(* Logix 5000 project; controller CIP vendor 1 type 14 code 106 rev 20.12; software revision 20.06; part 8 of 13 *)
(* tags used below, declared in another part *)
   MOA_OFF : DINT[10];
   MOA_ON : DINT[10];
   PV_Output_Status : INT[10];
   PV_Output_Status_IND : INT[10,16];
   PV_Status_Bit : BOOL;
   Time_Date : DINT[20];
(* MainProgram, continued *)

ROUTINE _10_PV_STATUS   (* ladder *)
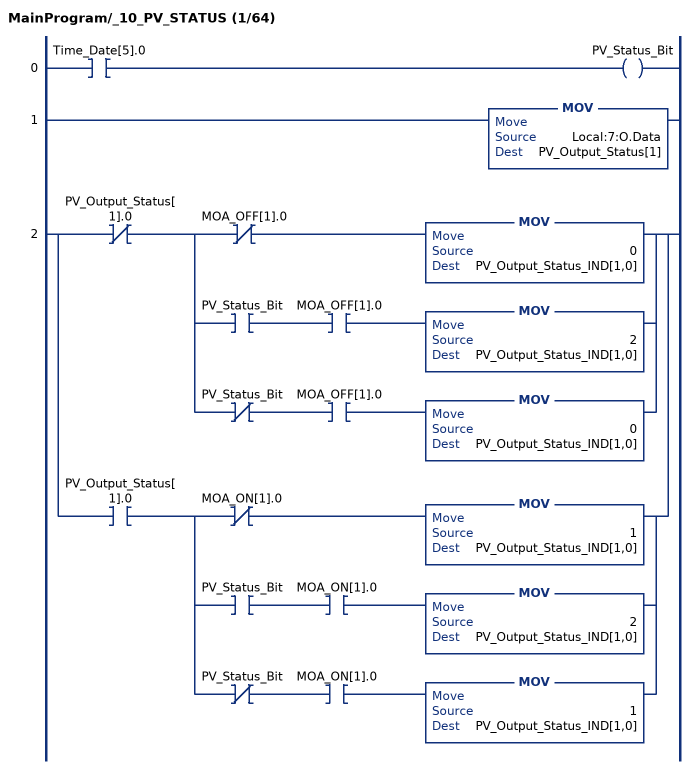
   0: XIC(Time_Date[5].0)OTE(PV_Status_Bit);
   1: MOV(Local:7:O.Data,PV_Output_Status[1]);
   2: [XIO(PV_Output_Status[1].0) [XIO(MOA_OFF[1].0) MOV(0,PV_Output_Status_IND[1,0]) ,XIC(PV_Status_Bit) XIC(MOA_OFF[1].0) MOV(2,PV_Output_Status_IND[1,0]) ,XIO(PV_Status_Bit) XIC(MOA_OFF[1].0) MOV(0,PV_Output_Status_IND[1,0]) ] ,XIC(PV_Output_Status[1].0) [XIO(MOA_ON[1].0) MOV(1,PV_Output_Status_IND[1,0]) ,XIC(PV_Status_Bit) XIC(MOA_ON[1].0) MOV(2,PV_Output_Status_IND[1,0]) ,XIO(PV_Status_Bit) XIC(MOA_ON[1].0) MOV(1,PV_Output_Status_IND[1,0]) ] ];
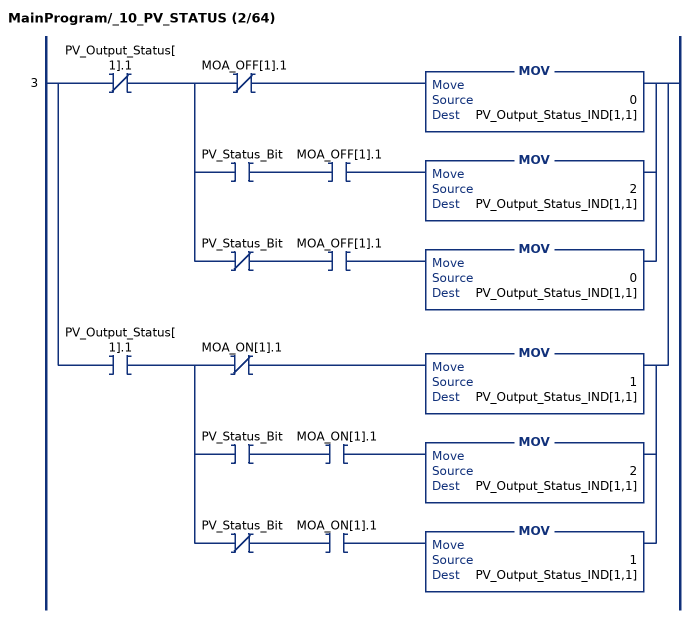
   3: [XIO(PV_Output_Status[1].1) [XIO(MOA_OFF[1].1) MOV(0,PV_Output_Status_IND[1,1]) ,XIC(PV_Status_Bit) XIC(MOA_OFF[1].1) MOV(2,PV_Output_Status_IND[1,1]) ,XIO(PV_Status_Bit) XIC(MOA_OFF[1].1) MOV(0,PV_Output_Status_IND[1,1]) ] ,XIC(PV_Output_Status[1].1) [XIO(MOA_ON[1].1) MOV(1,PV_Output_Status_IND[1,1]) ,XIC(PV_Status_Bit) XIC(MOA_ON[1].1) MOV(2,PV_Output_Status_IND[1,1]) ,XIO(PV_Status_Bit) XIC(MOA_ON[1].1) MOV(1,PV_Output_Status_IND[1,1]) ] ];
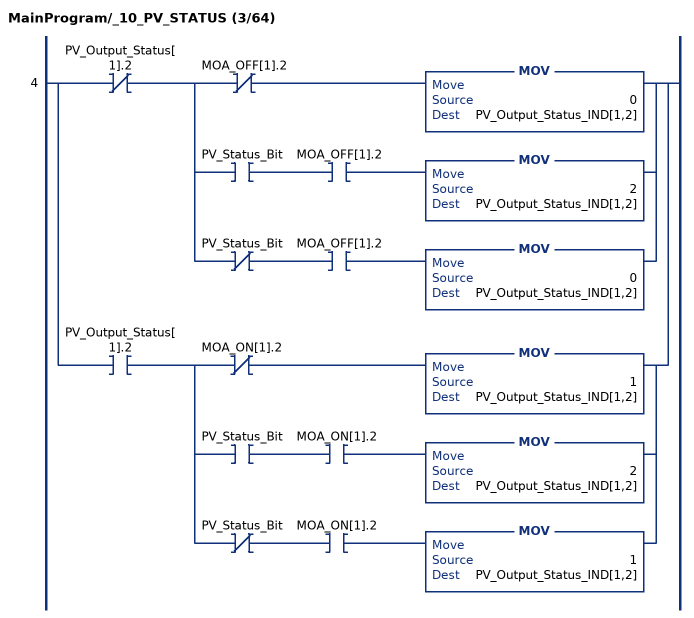
   4: [XIO(PV_Output_Status[1].2) [XIO(MOA_OFF[1].2) MOV(0,PV_Output_Status_IND[1,2]) ,XIC(PV_Status_Bit) XIC(MOA_OFF[1].2) MOV(2,PV_Output_Status_IND[1,2]) ,XIO(PV_Status_Bit) XIC(MOA_OFF[1].2) MOV(0,PV_Output_Status_IND[1,2]) ] ,XIC(PV_Output_Status[1].2) [XIO(MOA_ON[1].2) MOV(1,PV_Output_Status_IND[1,2]) ,XIC(PV_Status_Bit) XIC(MOA_ON[1].2) MOV(2,PV_Output_Status_IND[1,2]) ,XIO(PV_Status_Bit) XIC(MOA_ON[1].2) MOV(1,PV_Output_Status_IND[1,2]) ] ];
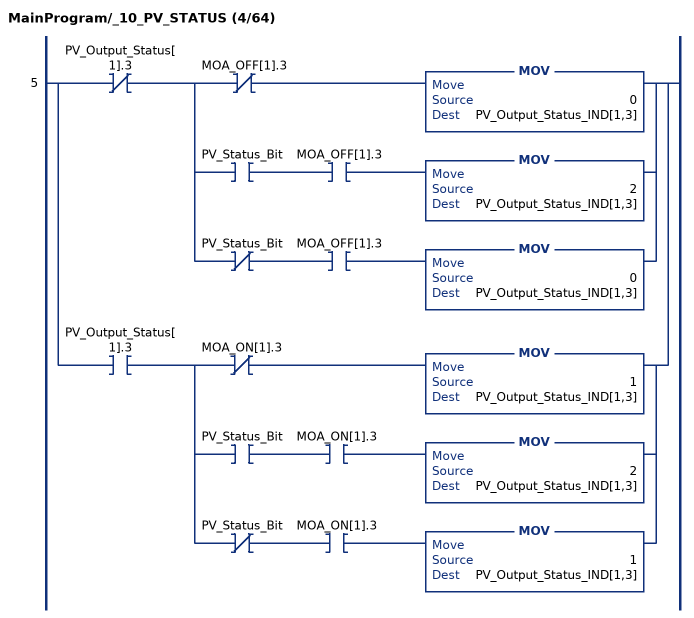
   5: [XIO(PV_Output_Status[1].3) [XIO(MOA_OFF[1].3) MOV(0,PV_Output_Status_IND[1,3]) ,XIC(PV_Status_Bit) XIC(MOA_OFF[1].3) MOV(2,PV_Output_Status_IND[1,3]) ,XIO(PV_Status_Bit) XIC(MOA_OFF[1].3) MOV(0,PV_Output_Status_IND[1,3]) ] ,XIC(PV_Output_Status[1].3) [XIO(MOA_ON[1].3) MOV(1,PV_Output_Status_IND[1,3]) ,XIC(PV_Status_Bit) XIC(MOA_ON[1].3) MOV(2,PV_Output_Status_IND[1,3]) ,XIO(PV_Status_Bit) XIC(MOA_ON[1].3) MOV(1,PV_Output_Status_IND[1,3]) ] ];
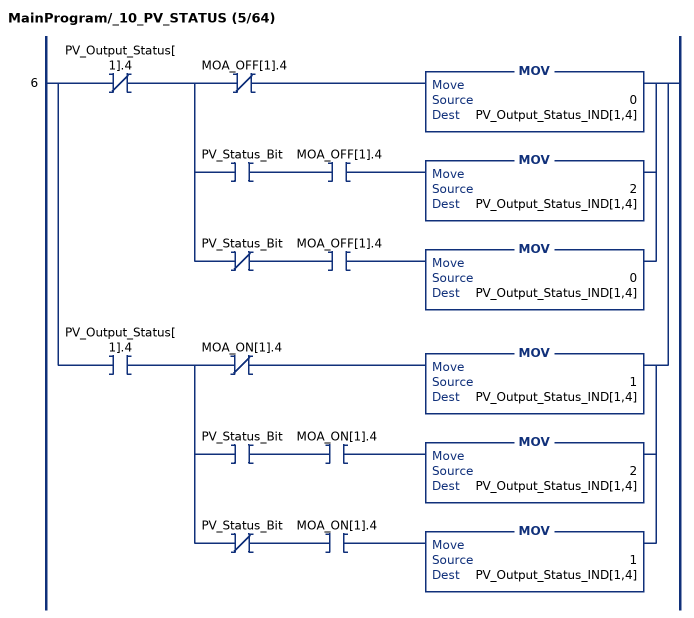
   6: [XIO(PV_Output_Status[1].4) [XIO(MOA_OFF[1].4) MOV(0,PV_Output_Status_IND[1,4]) ,XIC(PV_Status_Bit) XIC(MOA_OFF[1].4) MOV(2,PV_Output_Status_IND[1,4]) ,XIO(PV_Status_Bit) XIC(MOA_OFF[1].4) MOV(0,PV_Output_Status_IND[1,4]) ] ,XIC(PV_Output_Status[1].4) [XIO(MOA_ON[1].4) MOV(1,PV_Output_Status_IND[1,4]) ,XIC(PV_Status_Bit) XIC(MOA_ON[1].4) MOV(2,PV_Output_Status_IND[1,4]) ,XIO(PV_Status_Bit) XIC(MOA_ON[1].4) MOV(1,PV_Output_Status_IND[1,4]) ] ];
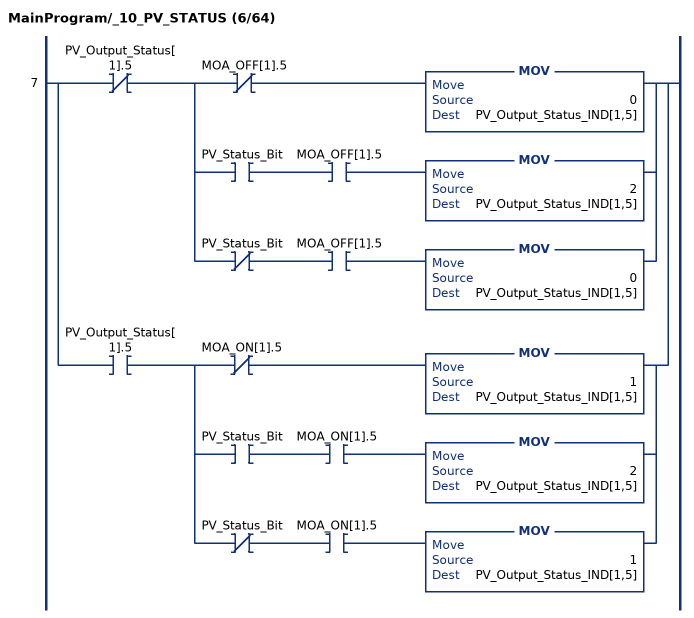
   7: [XIO(PV_Output_Status[1].5) [XIO(MOA_OFF[1].5) MOV(0,PV_Output_Status_IND[1,5]) ,XIC(PV_Status_Bit) XIC(MOA_OFF[1].5) MOV(2,PV_Output_Status_IND[1,5]) ,XIO(PV_Status_Bit) XIC(MOA_OFF[1].5) MOV(0,PV_Output_Status_IND[1,5]) ] ,XIC(PV_Output_Status[1].5) [XIO(MOA_ON[1].5) MOV(1,PV_Output_Status_IND[1,5]) ,XIC(PV_Status_Bit) XIC(MOA_ON[1].5) MOV(2,PV_Output_Status_IND[1,5]) ,XIO(PV_Status_Bit) XIC(MOA_ON[1].5) MOV(1,PV_Output_Status_IND[1,5]) ] ];
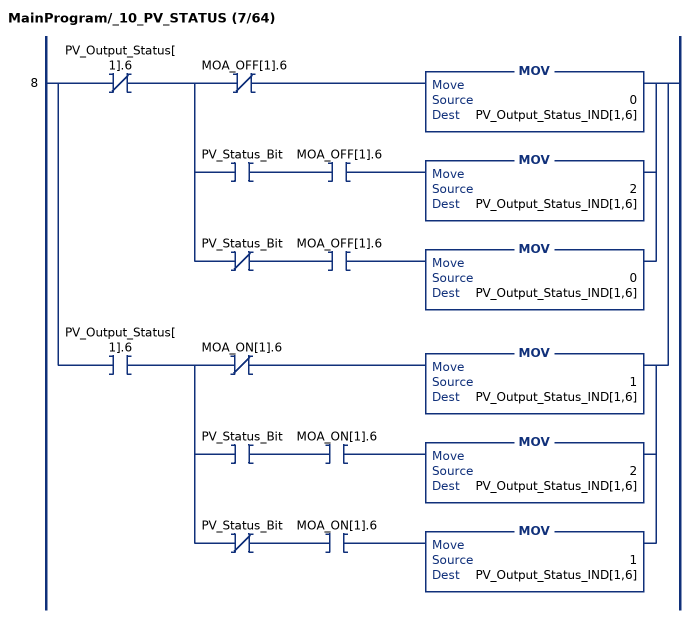
   8: [XIO(PV_Output_Status[1].6) [XIO(MOA_OFF[1].6) MOV(0,PV_Output_Status_IND[1,6]) ,XIC(PV_Status_Bit) XIC(MOA_OFF[1].6) MOV(2,PV_Output_Status_IND[1,6]) ,XIO(PV_Status_Bit) XIC(MOA_OFF[1].6) MOV(0,PV_Output_Status_IND[1,6]) ] ,XIC(PV_Output_Status[1].6) [XIO(MOA_ON[1].6) MOV(1,PV_Output_Status_IND[1,6]) ,XIC(PV_Status_Bit) XIC(MOA_ON[1].6) MOV(2,PV_Output_Status_IND[1,6]) ,XIO(PV_Status_Bit) XIC(MOA_ON[1].6) MOV(1,PV_Output_Status_IND[1,6]) ] ];
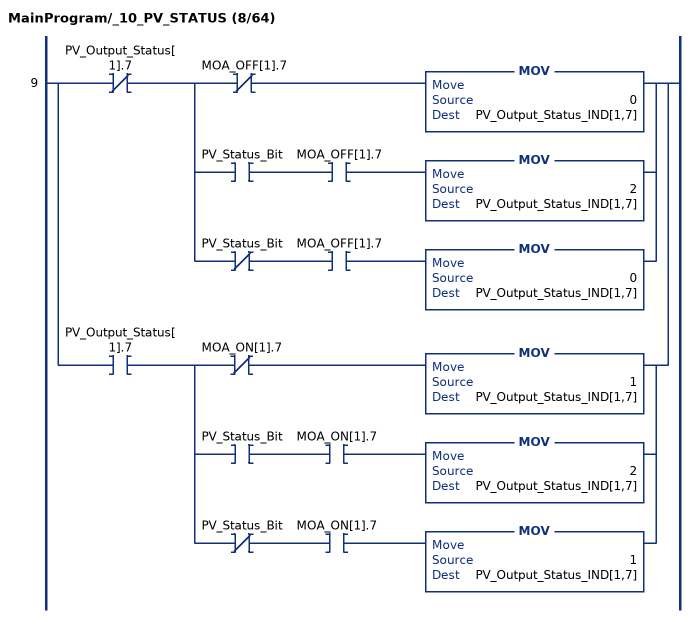
   9: [XIO(PV_Output_Status[1].7) [XIO(MOA_OFF[1].7) MOV(0,PV_Output_Status_IND[1,7]) ,XIC(PV_Status_Bit) XIC(MOA_OFF[1].7) MOV(2,PV_Output_Status_IND[1,7]) ,XIO(PV_Status_Bit) XIC(MOA_OFF[1].7) MOV(0,PV_Output_Status_IND[1,7]) ] ,XIC(PV_Output_Status[1].7) [XIO(MOA_ON[1].7) MOV(1,PV_Output_Status_IND[1,7]) ,XIC(PV_Status_Bit) XIC(MOA_ON[1].7) MOV(2,PV_Output_Status_IND[1,7]) ,XIO(PV_Status_Bit) XIC(MOA_ON[1].7) MOV(1,PV_Output_Status_IND[1,7]) ] ];
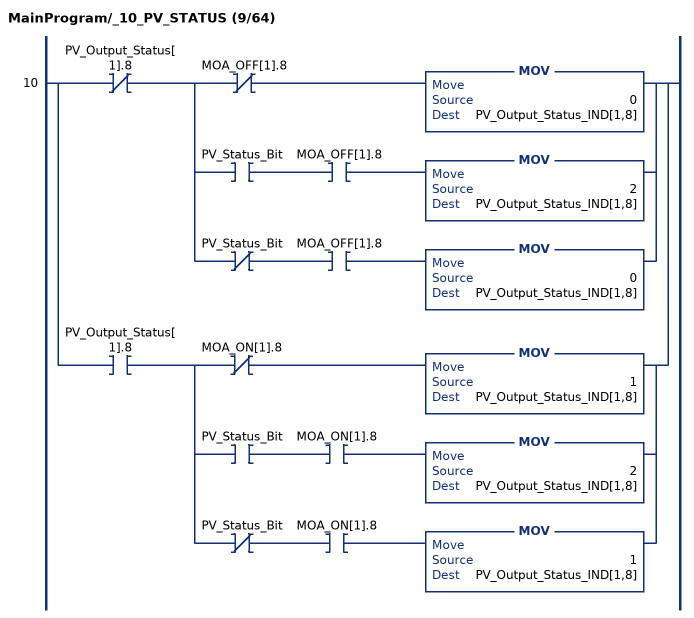
   10: [XIO(PV_Output_Status[1].8) [XIO(MOA_OFF[1].8) MOV(0,PV_Output_Status_IND[1,8]) ,XIC(PV_Status_Bit) XIC(MOA_OFF[1].8) MOV(2,PV_Output_Status_IND[1,8]) ,XIO(PV_Status_Bit) XIC(MOA_OFF[1].8) MOV(0,PV_Output_Status_IND[1,8]) ] ,XIC(PV_Output_Status[1].8) [XIO(MOA_ON[1].8) MOV(1,PV_Output_Status_IND[1,8]) ,XIC(PV_Status_Bit) XIC(MOA_ON[1].8) MOV(2,PV_Output_Status_IND[1,8]) ,XIO(PV_Status_Bit) XIC(MOA_ON[1].8) MOV(1,PV_Output_Status_IND[1,8]) ] ];
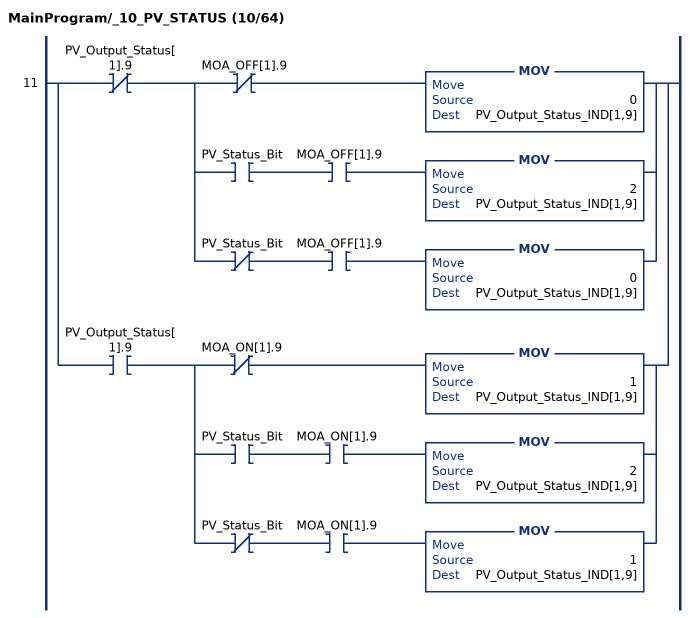
   11: [XIO(PV_Output_Status[1].9) [XIO(MOA_OFF[1].9) MOV(0,PV_Output_Status_IND[1,9]) ,XIC(PV_Status_Bit) XIC(MOA_OFF[1].9) MOV(2,PV_Output_Status_IND[1,9]) ,XIO(PV_Status_Bit) XIC(MOA_OFF[1].9) MOV(0,PV_Output_Status_IND[1,9]) ] ,XIC(PV_Output_Status[1].9) [XIO(MOA_ON[1].9) MOV(1,PV_Output_Status_IND[1,9]) ,XIC(PV_Status_Bit) XIC(MOA_ON[1].9) MOV(2,PV_Output_Status_IND[1,9]) ,XIO(PV_Status_Bit) XIC(MOA_ON[1].9) MOV(1,PV_Output_Status_IND[1,9]) ] ];
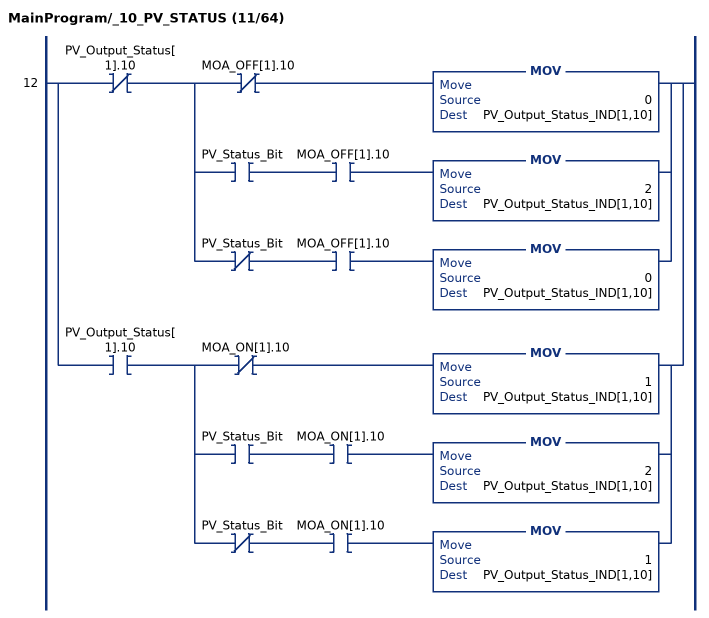
   12: [XIO(PV_Output_Status[1].10) [XIO(MOA_OFF[1].10) MOV(0,PV_Output_Status_IND[1,10]) ,XIC(PV_Status_Bit) XIC(MOA_OFF[1].10) MOV(2,PV_Output_Status_IND[1,10]) ,XIO(PV_Status_Bit) XIC(MOA_OFF[1].10) MOV(0,PV_Output_Status_IND[1,10]) ] ,XIC(PV_Output_Status[1].10) [XIO(MOA_ON[1].10) MOV(1,PV_Output_Status_IND[1,10]) ,XIC(PV_Status_Bit) XIC(MOA_ON[1].10) MOV(2,PV_Output_Status_IND[1,10]) ,XIO(PV_Status_Bit) XIC(MOA_ON[1].10) MOV(1,PV_Output_Status_IND[1,10]) ] ];
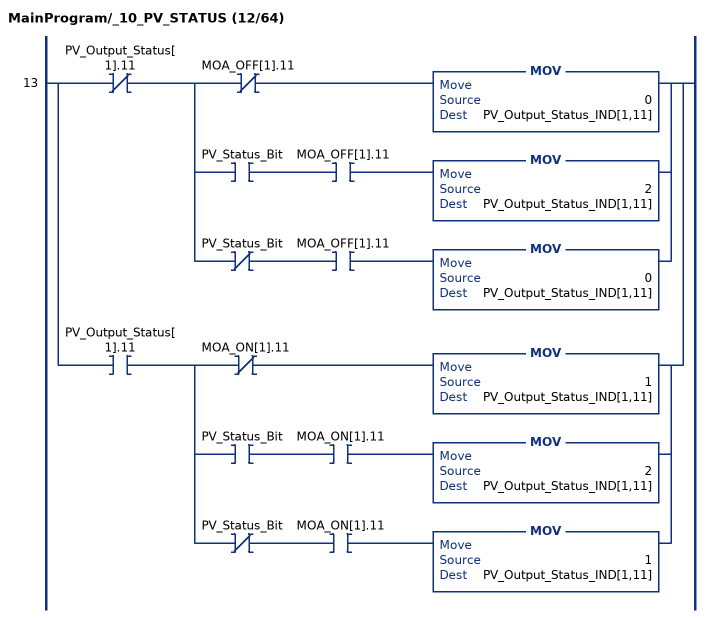
   13: [XIO(PV_Output_Status[1].11) [XIO(MOA_OFF[1].11) MOV(0,PV_Output_Status_IND[1,11]) ,XIC(PV_Status_Bit) XIC(MOA_OFF[1].11) MOV(2,PV_Output_Status_IND[1,11]) ,XIO(PV_Status_Bit) XIC(MOA_OFF[1].11) MOV(0,PV_Output_Status_IND[1,11]) ] ,XIC(PV_Output_Status[1].11) [XIO(MOA_ON[1].11) MOV(1,PV_Output_Status_IND[1,11]) ,XIC(PV_Status_Bit) XIC(MOA_ON[1].11) MOV(2,PV_Output_Status_IND[1,11]) ,XIO(PV_Status_Bit) XIC(MOA_ON[1].11) MOV(1,PV_Output_Status_IND[1,11]) ] ];
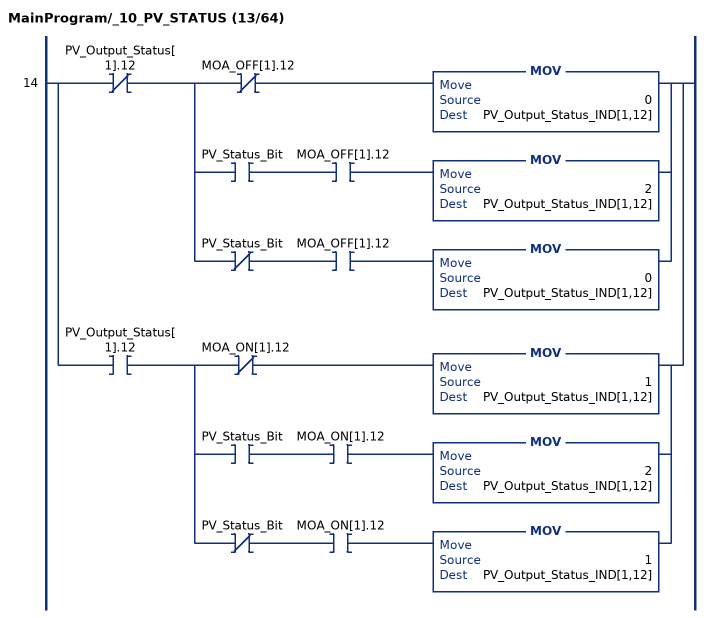
   14: [XIO(PV_Output_Status[1].12) [XIO(MOA_OFF[1].12) MOV(0,PV_Output_Status_IND[1,12]) ,XIC(PV_Status_Bit) XIC(MOA_OFF[1].12) MOV(2,PV_Output_Status_IND[1,12]) ,XIO(PV_Status_Bit) XIC(MOA_OFF[1].12) MOV(0,PV_Output_Status_IND[1,12]) ] ,XIC(PV_Output_Status[1].12) [XIO(MOA_ON[1].12) MOV(1,PV_Output_Status_IND[1,12]) ,XIC(PV_Status_Bit) XIC(MOA_ON[1].12) MOV(2,PV_Output_Status_IND[1,12]) ,XIO(PV_Status_Bit) XIC(MOA_ON[1].12) MOV(1,PV_Output_Status_IND[1,12]) ] ];
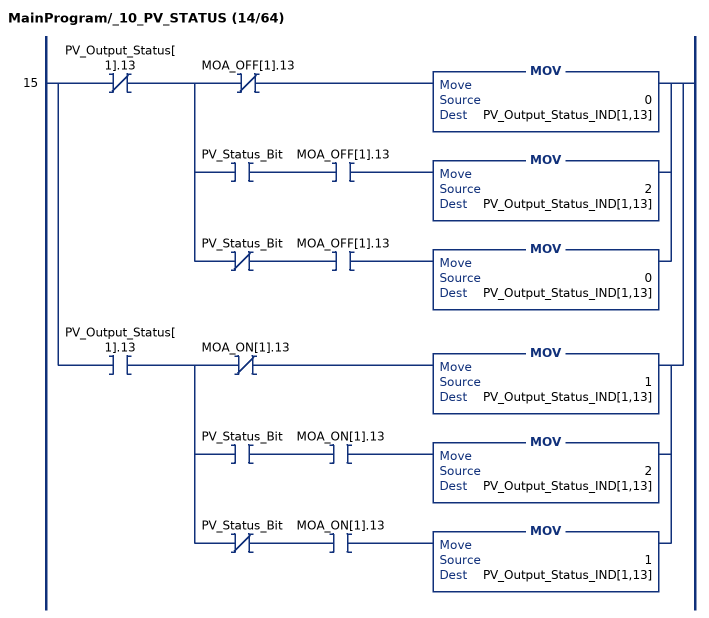
   15: [XIO(PV_Output_Status[1].13) [XIO(MOA_OFF[1].13) MOV(0,PV_Output_Status_IND[1,13]) ,XIC(PV_Status_Bit) XIC(MOA_OFF[1].13) MOV(2,PV_Output_Status_IND[1,13]) ,XIO(PV_Status_Bit) XIC(MOA_OFF[1].13) MOV(0,PV_Output_Status_IND[1,13]) ] ,XIC(PV_Output_Status[1].13) [XIO(MOA_ON[1].13) MOV(1,PV_Output_Status_IND[1,13]) ,XIC(PV_Status_Bit) XIC(MOA_ON[1].13) MOV(2,PV_Output_Status_IND[1,13]) ,XIO(PV_Status_Bit) XIC(MOA_ON[1].13) MOV(1,PV_Output_Status_IND[1,13]) ] ];
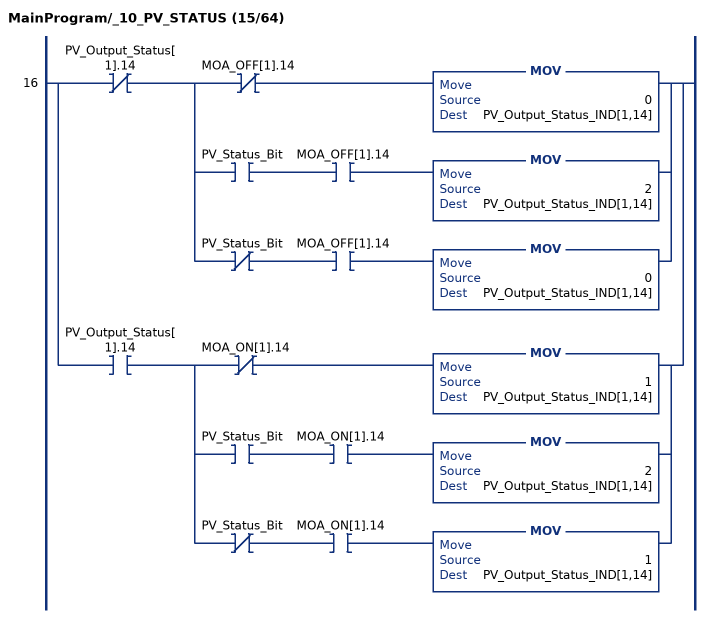
   16: [XIO(PV_Output_Status[1].14) [XIO(MOA_OFF[1].14) MOV(0,PV_Output_Status_IND[1,14]) ,XIC(PV_Status_Bit) XIC(MOA_OFF[1].14) MOV(2,PV_Output_Status_IND[1,14]) ,XIO(PV_Status_Bit) XIC(MOA_OFF[1].14) MOV(0,PV_Output_Status_IND[1,14]) ] ,XIC(PV_Output_Status[1].14) [XIO(MOA_ON[1].14) MOV(1,PV_Output_Status_IND[1,14]) ,XIC(PV_Status_Bit) XIC(MOA_ON[1].14) MOV(2,PV_Output_Status_IND[1,14]) ,XIO(PV_Status_Bit) XIC(MOA_ON[1].14) MOV(1,PV_Output_Status_IND[1,14]) ] ];
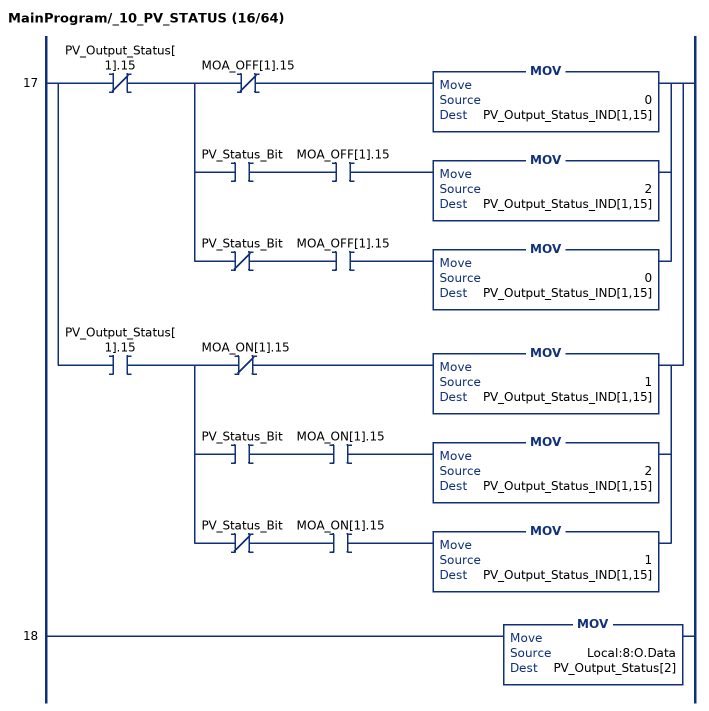
   17: [XIO(PV_Output_Status[1].15) [XIO(MOA_OFF[1].15) MOV(0,PV_Output_Status_IND[1,15]) ,XIC(PV_Status_Bit) XIC(MOA_OFF[1].15) MOV(2,PV_Output_Status_IND[1,15]) ,XIO(PV_Status_Bit) XIC(MOA_OFF[1].15) MOV(0,PV_Output_Status_IND[1,15]) ] ,XIC(PV_Output_Status[1].15) [XIO(MOA_ON[1].15) MOV(1,PV_Output_Status_IND[1,15]) ,XIC(PV_Status_Bit) XIC(MOA_ON[1].15) MOV(2,PV_Output_Status_IND[1,15]) ,XIO(PV_Status_Bit) XIC(MOA_ON[1].15) MOV(1,PV_Output_Status_IND[1,15]) ] ];
   18: MOV(Local:8:O.Data,PV_Output_Status[2]);
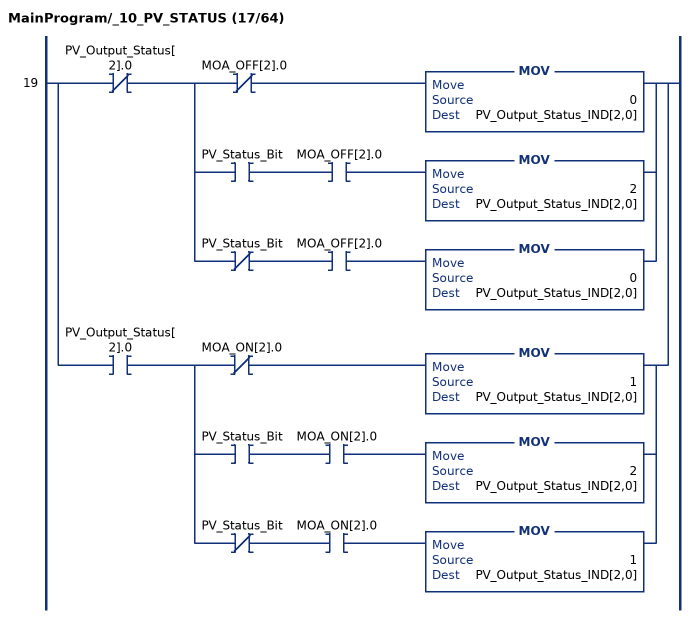
   19: [XIO(PV_Output_Status[2].0) [XIO(MOA_OFF[2].0) MOV(0,PV_Output_Status_IND[2,0]) ,XIC(PV_Status_Bit) XIC(MOA_OFF[2].0) MOV(2,PV_Output_Status_IND[2,0]) ,XIO(PV_Status_Bit) XIC(MOA_OFF[2].0) MOV(0,PV_Output_Status_IND[2,0]) ] ,XIC(PV_Output_Status[2].0) [XIO(MOA_ON[2].0) MOV(1,PV_Output_Status_IND[2,0]) ,XIC(PV_Status_Bit) XIC(MOA_ON[2].0) MOV(2,PV_Output_Status_IND[2,0]) ,XIO(PV_Status_Bit) XIC(MOA_ON[2].0) MOV(1,PV_Output_Status_IND[2,0]) ] ];
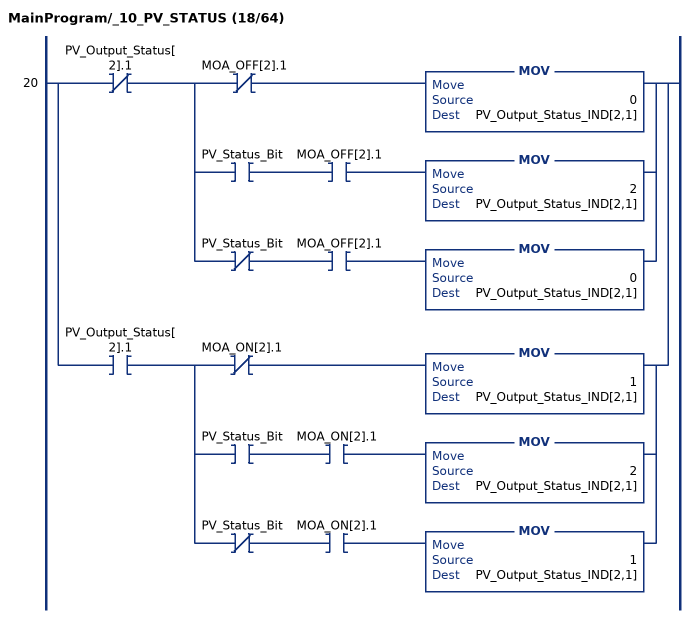
   20: [XIO(PV_Output_Status[2].1) [XIO(MOA_OFF[2].1) MOV(0,PV_Output_Status_IND[2,1]) ,XIC(PV_Status_Bit) XIC(MOA_OFF[2].1) MOV(2,PV_Output_Status_IND[2,1]) ,XIO(PV_Status_Bit) XIC(MOA_OFF[2].1) MOV(0,PV_Output_Status_IND[2,1]) ] ,XIC(PV_Output_Status[2].1) [XIO(MOA_ON[2].1) MOV(1,PV_Output_Status_IND[2,1]) ,XIC(PV_Status_Bit) XIC(MOA_ON[2].1) MOV(2,PV_Output_Status_IND[2,1]) ,XIO(PV_Status_Bit) XIC(MOA_ON[2].1) MOV(1,PV_Output_Status_IND[2,1]) ] ];
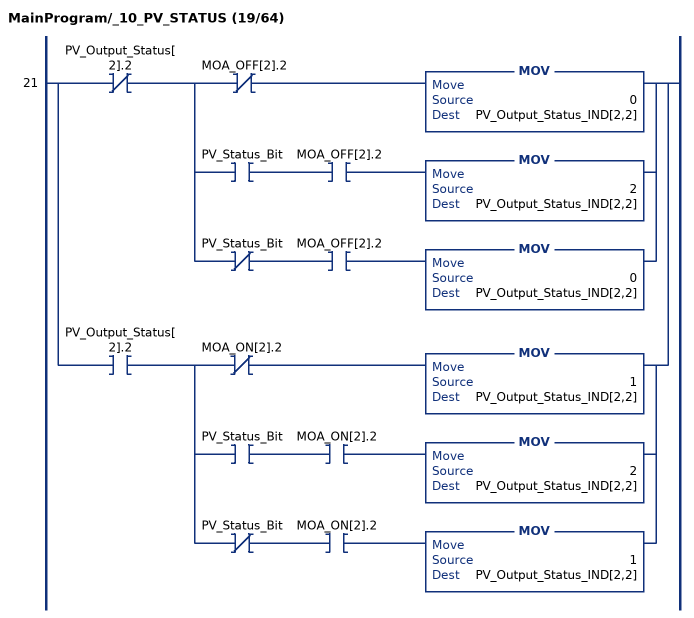
   21: [XIO(PV_Output_Status[2].2) [XIO(MOA_OFF[2].2) MOV(0,PV_Output_Status_IND[2,2]) ,XIC(PV_Status_Bit) XIC(MOA_OFF[2].2) MOV(2,PV_Output_Status_IND[2,2]) ,XIO(PV_Status_Bit) XIC(MOA_OFF[2].2) MOV(0,PV_Output_Status_IND[2,2]) ] ,XIC(PV_Output_Status[2].2) [XIO(MOA_ON[2].2) MOV(1,PV_Output_Status_IND[2,2]) ,XIC(PV_Status_Bit) XIC(MOA_ON[2].2) MOV(2,PV_Output_Status_IND[2,2]) ,XIO(PV_Status_Bit) XIC(MOA_ON[2].2) MOV(1,PV_Output_Status_IND[2,2]) ] ];
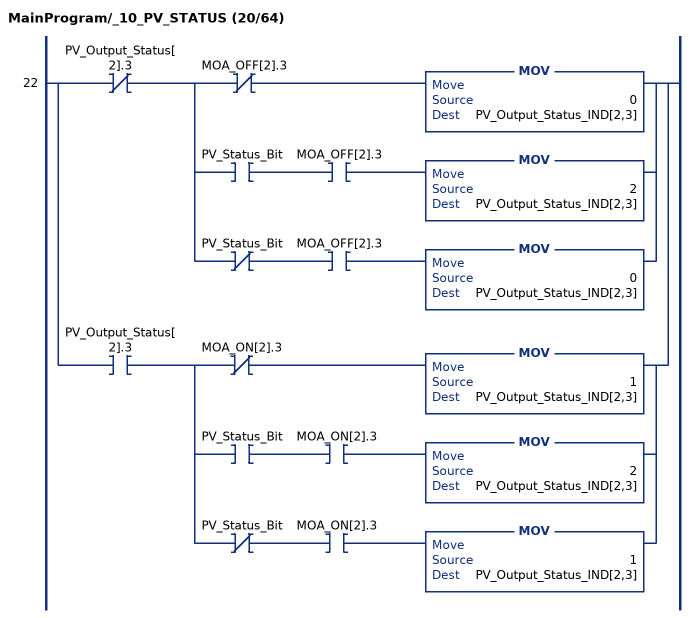
   22: [XIO(PV_Output_Status[2].3) [XIO(MOA_OFF[2].3) MOV(0,PV_Output_Status_IND[2,3]) ,XIC(PV_Status_Bit) XIC(MOA_OFF[2].3) MOV(2,PV_Output_Status_IND[2,3]) ,XIO(PV_Status_Bit) XIC(MOA_OFF[2].3) MOV(0,PV_Output_Status_IND[2,3]) ] ,XIC(PV_Output_Status[2].3) [XIO(MOA_ON[2].3) MOV(1,PV_Output_Status_IND[2,3]) ,XIC(PV_Status_Bit) XIC(MOA_ON[2].3) MOV(2,PV_Output_Status_IND[2,3]) ,XIO(PV_Status_Bit) XIC(MOA_ON[2].3) MOV(1,PV_Output_Status_IND[2,3]) ] ];
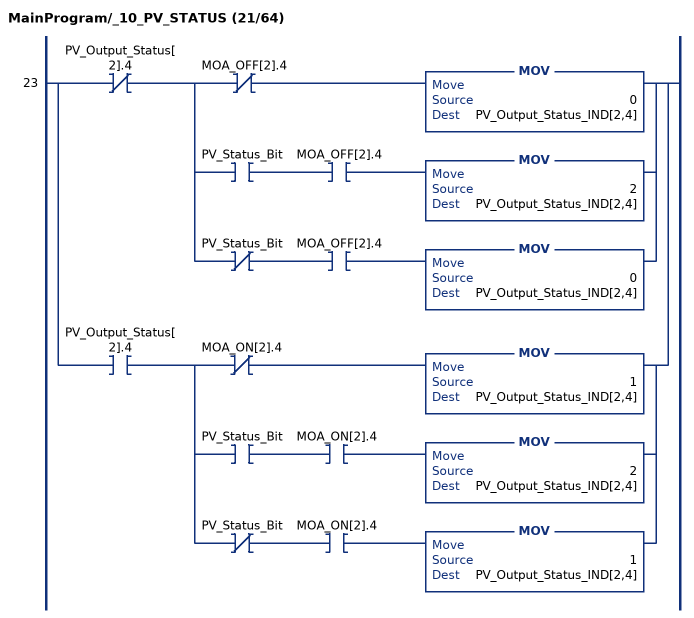
   23: [XIO(PV_Output_Status[2].4) [XIO(MOA_OFF[2].4) MOV(0,PV_Output_Status_IND[2,4]) ,XIC(PV_Status_Bit) XIC(MOA_OFF[2].4) MOV(2,PV_Output_Status_IND[2,4]) ,XIO(PV_Status_Bit) XIC(MOA_OFF[2].4) MOV(0,PV_Output_Status_IND[2,4]) ] ,XIC(PV_Output_Status[2].4) [XIO(MOA_ON[2].4) MOV(1,PV_Output_Status_IND[2,4]) ,XIC(PV_Status_Bit) XIC(MOA_ON[2].4) MOV(2,PV_Output_Status_IND[2,4]) ,XIO(PV_Status_Bit) XIC(MOA_ON[2].4) MOV(1,PV_Output_Status_IND[2,4]) ] ];
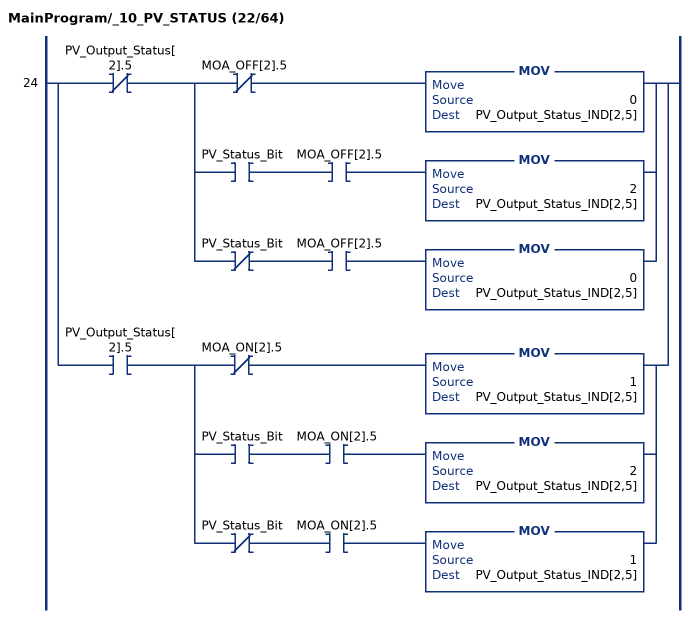
   24: [XIO(PV_Output_Status[2].5) [XIO(MOA_OFF[2].5) MOV(0,PV_Output_Status_IND[2,5]) ,XIC(PV_Status_Bit) XIC(MOA_OFF[2].5) MOV(2,PV_Output_Status_IND[2,5]) ,XIO(PV_Status_Bit) XIC(MOA_OFF[2].5) MOV(0,PV_Output_Status_IND[2,5]) ] ,XIC(PV_Output_Status[2].5) [XIO(MOA_ON[2].5) MOV(1,PV_Output_Status_IND[2,5]) ,XIC(PV_Status_Bit) XIC(MOA_ON[2].5) MOV(2,PV_Output_Status_IND[2,5]) ,XIO(PV_Status_Bit) XIC(MOA_ON[2].5) MOV(1,PV_Output_Status_IND[2,5]) ] ];
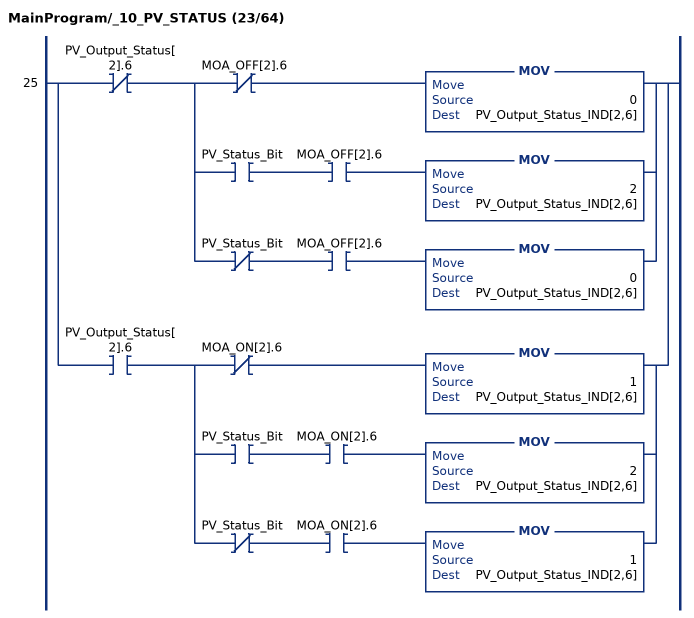
   25: [XIO(PV_Output_Status[2].6) [XIO(MOA_OFF[2].6) MOV(0,PV_Output_Status_IND[2,6]) ,XIC(PV_Status_Bit) XIC(MOA_OFF[2].6) MOV(2,PV_Output_Status_IND[2,6]) ,XIO(PV_Status_Bit) XIC(MOA_OFF[2].6) MOV(0,PV_Output_Status_IND[2,6]) ] ,XIC(PV_Output_Status[2].6) [XIO(MOA_ON[2].6) MOV(1,PV_Output_Status_IND[2,6]) ,XIC(PV_Status_Bit) XIC(MOA_ON[2].6) MOV(2,PV_Output_Status_IND[2,6]) ,XIO(PV_Status_Bit) XIC(MOA_ON[2].6) MOV(1,PV_Output_Status_IND[2,6]) ] ];
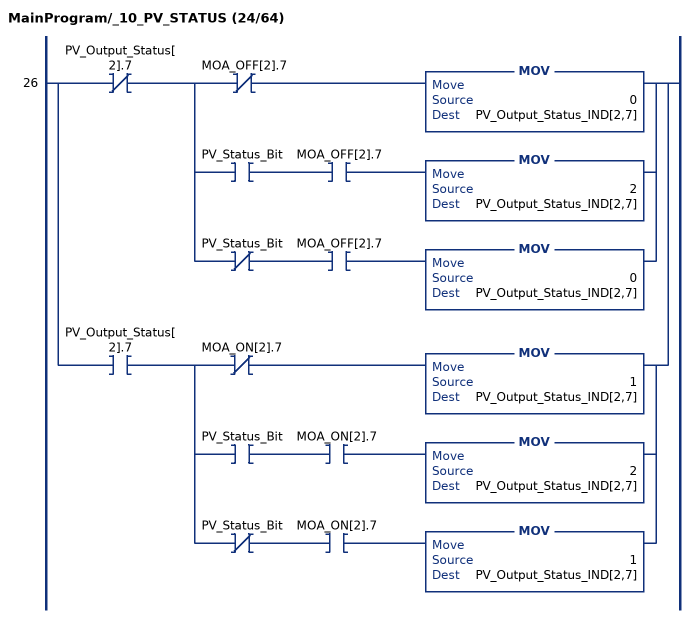
   26: [XIO(PV_Output_Status[2].7) [XIO(MOA_OFF[2].7) MOV(0,PV_Output_Status_IND[2,7]) ,XIC(PV_Status_Bit) XIC(MOA_OFF[2].7) MOV(2,PV_Output_Status_IND[2,7]) ,XIO(PV_Status_Bit) XIC(MOA_OFF[2].7) MOV(0,PV_Output_Status_IND[2,7]) ] ,XIC(PV_Output_Status[2].7) [XIO(MOA_ON[2].7) MOV(1,PV_Output_Status_IND[2,7]) ,XIC(PV_Status_Bit) XIC(MOA_ON[2].7) MOV(2,PV_Output_Status_IND[2,7]) ,XIO(PV_Status_Bit) XIC(MOA_ON[2].7) MOV(1,PV_Output_Status_IND[2,7]) ] ];
